(* IEC 61131-3 sources: llm-plc-st-eval/data/definitivo/gpt-4o-2024-08-06/I5/zero_shot, 3 files *)

(* ---- ejec_1.st ---- *)
```pascal
FUNCTION_BLOCK FB_Clasificadora
VAR_INPUT
    sensorPresencia : BOOL; // Sensor que detecta la presencia de una pieza
    sensorAltura : BOOL;    // Sensor que detecta si la pieza es alta
END_VAR

VAR_OUTPUT
    banda : BOOL;   // Salida para activar la banda transportadora
    piston : BOOL;  // Salida para activar el pistón desviador
    nAltas : INT;   // Contador de piezas altas
    nBajas : INT;   // Contador de piezas bajas
END_VAR

VAR
    timerRetraso : TON; // Temporizador para el retraso de 2 segundos
    timerPiston : TON;  // Temporizador para la activación del pistón durante 1 segundo
    piezaDetectada : BOOL; // Indica si una pieza ha sido detectada
    piezaAlta : BOOL; // Indica si la pieza detectada es alta
END_VAR

// Inicialización de la banda transportadora
banda := TRUE;

// Detección de una pieza
IF sensorPresencia AND NOT piezaDetectada THEN
    piezaDetectada := TRUE;
    piezaAlta := sensorAltura;
    timerRetraso(IN := TRUE, PT := T#2S); // Inicia el temporizador de retraso
END_IF

// Manejo del temporizador de retraso
IF timerRetraso.Q THEN
    timerRetraso(IN := FALSE); // Detiene el temporizador de retraso

    IF piezaAlta THEN
        timerPiston(IN := TRUE, PT := T#1S); // Inicia el temporizador del pistón
        nAltas := nAltas + 1; // Incrementa el contador de piezas altas
    ELSE
        nBajas := nBajas + 1; // Incrementa el contador de piezas bajas
    END_IF

    piezaDetectada := FALSE; // Reinicia la detección de pieza
END_IF

// Manejo del temporizador del pistón
IF timerPiston.Q THEN
    piston := FALSE; // Desactiva el pistón
    timerPiston(IN := FALSE); // Detiene el temporizador del pistón
ELSE
    piston := timerPiston.Q; // Activa el pistón mientras el temporizador está activo
END_IF

END_FUNCTION_BLOCK
```

Este código implementa un bloque de función `FB_Clasificadora` que controla una banda transportadora clasificadora. La banda funciona continuamente, y las piezas se clasifican en altas y bajas según la entrada de los sensores. El pistón se activa para desviar las piezas altas después de un retraso de 2 segundos y se mantiene activo durante 1 segundo. Los contadores `nAltas` y `nBajas` llevan un registro del número de piezas altas y bajas, respectivamente.

(* ---- ejec_2.st ---- *)
```pascal
FUNCTION_BLOCK FB_Clasificadora
VAR_INPUT
    sensorPresencia : BOOL; // Sensor que detecta la presencia de una pieza
    sensorAltura : BOOL;    // Sensor que detecta si la pieza es alta
END_VAR

VAR_OUTPUT
    banda : BOOL := TRUE;   // Salida que activa la banda transportadora
    piston : BOOL := FALSE; // Salida que activa el pistón desviador
    nAltas : INT := 0;      // Contador de piezas altas
    nBajas : INT := 0;      // Contador de piezas bajas
END_VAR

VAR
    estadoAnteriorPresencia : BOOL := FALSE; // Estado anterior del sensor de presencia
    temporizadorRetraso : TON;              // Temporizador para el retraso de 2 segundos
    temporizadorPiston : TON;               // Temporizador para la duración de 1 segundo del pistón
    activarPiston : BOOL := FALSE;          // Bandera para activar el pistón
END_VAR

// Inicialización de los temporizadores
temporizadorRetraso(IN := FALSE, PT := T#2S);
temporizadorPiston(IN := FALSE, PT := T#1S);

// Detectar flanco de subida del sensor de presencia
IF (sensorPresencia AND NOT estadoAnteriorPresencia) THEN
    IF sensorAltura THEN
        // Iniciar temporizador de retraso para piezas altas
        temporizadorRetraso(IN := TRUE);
        activarPiston := TRUE;
    ELSE
        // Incrementar contador de piezas bajas
        nBajas := nBajas + 1;
    END_IF;
END_IF;

// Actualizar estado anterior del sensor de presencia
estadoAnteriorPresencia := sensorPresencia;

// Control del pistón
IF activarPiston THEN
    // Si el temporizador de retraso ha terminado, iniciar temporizador del pistón
    IF temporizadorRetraso.Q THEN
        temporizadorPiston(IN := TRUE);
        temporizadorRetraso(IN := FALSE);
    END_IF;

    // Activar el pistón durante 1 segundo
    IF temporizadorPiston.Q THEN
        piston := FALSE;
        temporizadorPiston(IN := FALSE);
        activarPiston := FALSE;
        nAltas := nAltas + 1; // Incrementar contador de piezas altas
    ELSE
        piston := TRUE;
    END_IF;
ELSE
    piston := FALSE;
END_IF;

banda := TRUE; // La banda siempre está activa
END_FUNCTION_BLOCK
```

(* ---- ejec_3.st ---- *)
```pascal
FUNCTION_BLOCK FB_Clasificadora
VAR_INPUT
    sensorPresencia : BOOL;  // Sensor que detecta la presencia de una pieza
    sensorAltura : BOOL;     // Sensor que detecta si la pieza es alta
END_VAR

VAR_OUTPUT
    banda : BOOL;            // Salida para activar la banda transportadora
    piston : BOOL;           // Salida para activar el pistón desviador
    nAltas : INT;            // Contador de piezas altas
    nBajas : INT;            // Contador de piezas bajas
END_VAR

VAR
    timerRetraso : TON;      // Temporizador para retrasar la activación del pistón
    timerDuracion : TON;     // Temporizador para la duración del pistón activado
    presenciaDetectada : BOOL; // Indica si se ha detectado una pieza
    piezaAlta : BOOL;        // Indica si la pieza detectada es alta
END_VAR

// Inicialización de la banda transportadora
banda := TRUE;

// Detección de una pieza
IF sensorPresencia AND NOT presenciaDetectada THEN
    presenciaDetectada := TRUE;
    piezaAlta := sensorAltura;

    // Iniciar temporizador de retraso si la pieza es alta
    IF piezaAlta THEN
        timerRetraso(IN := TRUE, PT := T#2S);
    ELSE
        nBajas := nBajas + 1; // Incrementar contador de piezas bajas
    END_IF
END_IF

// Manejo del temporizador de retraso
IF timerRetraso.Q THEN
    timerRetraso(IN := FALSE);
    timerDuracion(IN := TRUE, PT := T#1S);
    piston := TRUE;
END_IF

// Manejo del temporizador de duración del pistón
IF timerDuracion.Q THEN
    timerDuracion(IN := FALSE);
    piston := FALSE;
    nAltas := nAltas + 1; // Incrementar contador de piezas altas
END_IF

// Reiniciar detección de presencia
IF NOT sensorPresencia THEN
    presenciaDetectada := FALSE;
END_IF

END_FUNCTION_BLOCK
```

Este código implementa un bloque de función para controlar una banda transportadora clasificadora. La banda está siempre activa, y el pistón se activa para desviar piezas altas después de un retraso de 2 segundos, permaneciendo activo durante 1 segundo. Las piezas altas y bajas se cuentan en `nAltas` y `nBajas`, respectivamente.
